Fanuc KAREL source: KC00048.KL

PROGRAM KC00048
%NOLOCKGROUP
%ENVIRONMENT REGOPE
VAR
  I: INTEGER
  J: INTEGER
  K: INTEGER
  R: REAL
  B: BOOLEAN
  S: STRING[80]
  T: STRING[80]
  P: PATH
  Q: PATH
  AI: ARRAY[8] OF INTEGER
  AB: ARRAY[244] OF BYTE
  EP: XYZWPREXT
BEGIN
  SET_TPE_EPOS_REG(I,EP,J)
END KC00048
